// TIA Portal project "ifm-O3D3xx_S7-1200_V16" (V16)

(* hardware
DEVICE "S7-1200 station_1"  S7-1200 Station
   slot 0: "Rack_0"  S7-1200 Rack  Rack  V1.0
   slot 1: "PLC_1"  CPU 1212C AC/DC/Rly  6ES7 212-1BE40-0XB0  V4.4
DEVICE "GSD device_1"  GSD.Device.PN
   slot 0: "Rack"  Rack  V1.0
   slot 0: "O3D3xx"  O3D3XX-PN  O3D3xx  Z1.0
      slot 0: "Standard"  Standard
      slot 1: "Interface"  Interface
         slot 1: "RJ45 10/100 MBit/s"  RJ45 10/100 MBit/s
   slot 1: "450 bytes I_1"  450 bytes I  1.0
      slot 0: "450 bytes I"  450 bytes I
   slot 2: "8 bytes O_1"  8 bytes O  1.0
      slot 0: "8 bytes O"  8 bytes O
DEVICE "HMI_1"  TP700 Comfort
   slot 0: "HMI_1"  TP700 Comfort  6AV2 124-0GC01-0AX0  16.0.0.0
   slot 1: "HMI_RT_1"  TP700 Comfort  6AV2 124-0GC01-0AX0  16.0.0.0
   slot 5: "HMI_1.IE_CP_1"  PROFINET Interface  16.0.0.0
      slot 1: "PROFINET Interface_1"  PROFINET Interface
         slot 1: "Port_1"  Port
         slot 2: "Port_2"  Port
   slot 7: "HMI_1.MPI/DP_CP_1"  MPI/DP Interface  16.0.0.0
DEVICE "GSD device_2"  GSD.Device.PN
   slot 0: "Rack"  Rack  V1.0
   slot 0: "AL1100"  AL1100  AL1100
      slot 0: "AL1100"  AL1100
      slot 1: "X1"  X1
         slot 1: "Port 1"  Port 1
         slot 2: "Port 2"  Port 2
   slot 1: "4 Ports_1"  4 Ports  AL1100
      slot 0: "IO-Link Master"  IO-Link Master
   slot 1: "IO-Link In/Out 32/32 Byte + PQI"  IO-Link In/Out 32/32 Byte + PQI
*)

// ===== PLC "PLC_1"  CPU 1212C AC/DC/Rly =====

VAR_GLOBAL   // PLC tag table "Default tag table"
   "Trigger" AT %M0.0 : Bool;
   "AppNo" AT %MW2 : UInt;
   "GetCounters" AT %M0.1 : Bool;
   "ScrapRate" AT %MD6 : UDInt;
   "Scrap_Alarm" AT %M0.2 : Bool;
   "My_Row_is_OK" AT %M0.3 : Bool;
   "Big Box" AT %M0.4 : Bool;
   "Tag present" AT %I519.2 : Bool;
   "TagValue" AT %IB520 : Byte;
END_VAR

DATA_BLOCK "O3D3xx_Trigger_DB"   // DB1
{ S7_Optimized_Access := 'TRUE' }
AUTHOR : ifm-sy-tl
FAMILY : O3D3xx
VERSION : 1.0
// stored: InstanceOfName O3D3xx_Trigger
"O3D3xx_Trigger"
BEGIN
END_DATA_BLOCK

DATA_BLOCK "O3D3xx_Dimensioning_DB"   // DB2
{ S7_Optimized_Access := 'TRUE' }
AUTHOR : ifm-sy-tl
FAMILY : O3D3xx
VERSION : 1.0
// stored: InstanceOfName O3D3xx_Dimensioning
"O3D3xx_Dimensioning"
BEGIN
END_DATA_BLOCK

DATA_BLOCK "O3D3xx_Completeness_DB"   // DB3
{ S7_Optimized_Access := 'TRUE' }
AUTHOR : ifm-sy-tl
FAMILY : O3D3xx
VERSION : 1.0
// stored: InstanceOfName O3D3xx_Completeness
"O3D3xx_Completeness"
BEGIN
END_DATA_BLOCK

DATA_BLOCK "O3D3xx_GetStatistics_DB"   // DB4
{ S7_Optimized_Access := 'TRUE' }
AUTHOR : ifm-sy-tl
FAMILY : O3D3xx
VERSION : 1.0
// stored: InstanceOfName O3D3xx_GetStatistics
"O3D3xx_GetStatistics"
BEGIN
END_DATA_BLOCK

DATA_BLOCK "ReadData"   // DB5
{ S7_Optimized_Access := 'TRUE' }
VERSION : 0.1
   VAR
      RFIDValue : Byte;
      Object : Struct
         Length : Int;
         Width : Int;
         Height : Int;
      END_STRUCT;
   END_VAR
BEGIN
END_DATA_BLOCK

FUNCTION_BLOCK "O3D3xx_GetStatistics"   // FB8, SCL
TITLE = Get Statistics
{ S7_Optimized_Access := 'TRUE' }
AUTHOR : ifm-sy-tl
FAMILY : O3D3xx
VERSION : 1.1
// executes a "Get Statistics" command and provides the statistics of total, pass and fail readings
   VAR_INPUT
      HW_ID : Hw_Device;   // hardware identifier of the O3D3xx sensor
      Execute : Bool;   // execute Get Statistics command
      TimeoutTime : Time := T#500ms;   // timeout time
   END_VAR
   VAR_OUTPUT
      Done : Bool;   // completed without error
      Busy : Bool;   // command in process
      Error : Bool;   // error occurred
      Status : Word;   // status or error code
      CmdErrorCode : UDInt;   // command error code from O3D3xx sensor
      SysErrorCode : UDInt;   // system error code from O3D3xx sensor
      Total : UDInt;   // total readings
      Pass : UDInt;   // passed readings
      Fail : UDInt;   // failed readings
   END_VAR
   VAR
      tonTimeout : TON_TIME;   // timeout timer of command processing
      diCmdErrorCode : UDInt;   // command error code from O3D3xx sensor
      diSysErrorCode : UDInt;   // system error code from O3D3xx sensor
      wErrorCode : Word;   // current error code of the FB
      iState : Int;   // state of the state machine
      diTotal : UDInt;   // total readings
      diPass : UDInt;   // passed readings
      diFail : UDInt;   // failed readings
   END_VAR
   VAR_TEMP
      Addr : GEOADDR;   // GEO address of the module
      HWModuleID : Hw_Io;   // hardware ID the data module
      DIModuleInAddr : UDInt;   // input address of O3D3xx data
      DIModuleOutAddr : UDInt;   // output address of O3D3xx data
      DIDummy : UDInt;   // dummy
      IModuleInLength : UInt;   // size of data from O3D3xx
      IModuleOutLength : UInt;   // size of data to O3D3xx
      IDummy : UInt;   // dummy
      WCmd : Word;   // command word
      WMirror : Word;   // mirror word
      IResult : Int;   // result of system function
      XDone : Bool;   // task completed
      XError : Bool;   // error detected
      XErrorHW : Bool;   // error hardware assignment
   END_VAR
   VAR CONSTANT
      StateIdle : Int := 16#7000;   // state machine "idle"
      StateSensorRdy : Int := 16#7001;   // state machine "sensor ready"
      StateDeleteError : Int := 16#7002;   // state machine "delete error bit"
      StateGetStatistics : Int := 16#7801;   // state machine "get statistics"
      StateGetError : Int := 16#7601;   // state machine "get error code"
      StateDone : Int := 16#0000;   // state machine "completed"
      StateError : Int := 16#FFFF;   // state machine "error occurred"
   END_VAR
BEGIN
   // Sample program for reading the statistics from an ifm O3D3xx sensor
   // connected to the PLC as Profinet-IO device

   // Function Block Version 1.1.00

   // Description:
   (*
   This FB can be used with an ifm O3D3xx sensor that is connected as Profinet-IO device.
   The core of this FB is to execute a Get Statistics command.
   *)
   // ******************************************************************************************************
   // Disclaimer OF Warranties
   (*
   ifm disclaims to the fullest extent authorized by law any and all warranties,
   whether express or implied, including, without limitation,
   any implied warranties of title, non-infringement, quiet enjoyment,
   integration, merchantability or fitness for a particular purpose.

   Without limitation of the foregoing, ifm expressly does not warrant that:
   (a)  the software will meet your requirements or expectations;
   (b)  the software or the software content will be free of bugs, errors,
        viruses or other defects;
   (c)  any results, output, or data provided through or generated by the software
        will be accurate, up-to-date, complete or reliable;
   (d)  the software will be compatible with third party software;
   (e)  any errors in the software will be corrected


   DEMO SOFTWARE AND TEMPLATES

   Demo software and templates are provided “as is” and “as available”,
   without any warranty of any kind, either express or implied.
   The User acknowledges and agrees to use the software at User’s own risk.
   In no event shall ifm be held liable for any direct, indirect, incidental
   or consequential damages arising out of the use of or inability to use the software.
   User may use the software solely for demonstration purposes
   and to assess the software functionalities and capabilities.


   Software written specifically for Customer

   1. The software created and used is put together by ifm specially to the customer
      using modular software components made by ifm for numerous applications (Standard software modules)
      and adapted to the contractual service required (customer-specific application program).

   2. Upon complete payment of the purchase price for the customer-specific application program,
      ifm transfers the non-exclusive, locally and temporarily unrestricted usage right
      thereof to the customer, without the customer acquiring any rights of any kind
      to the standard software module on which the individual or customer-specific adaptation is based.
      Notwithstanding these provisions, ifm reserves the right to produce and offer
      customer specific software solutions of the same kind for other customers
      based on other terms of reference. In any case ifm retains a simple right of usage
      of the customer–specific solution for internal purposes.

   3. Upon acceptance of the program, User acknowledges and agrees to use the software
      at User’s own risk. User also acknowledges and agrees upon acceptance of the program
      that the software meets the requirements of the specifications agreed upon.
      ifm disclaims any and all warranties, in particular regarding fitness of the software
      for a particular purpose.
   ******************************************************************************************************
   *)

   REGION get addresses and size of O3D3xx data

     // read GEO address of O3D3xx sensor
     #IResult := LOG2GEO(LADDR := #HW_ID, GEOADDR := #Addr);
     #XErrorHW := #IResult <> 0 OR #Addr.AREA <> 1;  // check for error and AREA = PROFINET IO

     #Addr.HWTYPE := 4;  // set hardware type = Module
     #Addr.SUBSLOT := 0;  // set subslot

     REGION  get address and size of INPUT data from O3D3xx
       IF NOT #XErrorHW THEN
         #Addr.SLOT := 1;  // set slot = 1 (slot of INPUT data in O3D3xx configuration)
         #IResult := GEO2LOG(GEOADDR := #Addr, LADDR => #HWModuleID);  // get HW_ID of INPUT data module
         #XErrorHW := #IResult <> 0;  // check for error
       END_IF;
       IF NOT #XErrorHW THEN
         // get IO address of INPUT data
         #IResult := RD_ADDR(LADDR := #HWModuleID,
                             PIADDR => #DIModuleInAddr,
                             PICount => #IModuleInLength,
                             PQADDR => #DIDummy,
                             PQCount => #IDummy);
         #XErrorHW := #IResult <> 0 OR #IDummy <> 0 OR #IModuleInLength <> 64 AND #IModuleInLength <> 450;  // check for error and check size
       END_IF;
     END_REGION get address and size of INPUT data from O3D3xx

     REGION get address and size of OUTPUT data to O3D3xx
       IF NOT #XErrorHW THEN
         #Addr.SLOT := 2;  // set slot = 2 (slot of OUTPUT data in O3D3xx configuration)
         #IResult := GEO2LOG(GEOADDR := #Addr, LADDR => #HWModuleID);  // get HW_ID of OUTPUT data module
         #XErrorHW := #IResult <> 0;  // check for error
       END_IF;
       IF NOT #XErrorHW THEN
         // get IO address of OUTPUT data
         #IResult := RD_ADDR(LADDR := #HWModuleID,
                             PIADDR => #DIDummy,
                             PICount => #IDummy,
                             PQADDR => #DIModuleOutAddr,
                             PQCount => #IModuleOutLength);
         #XErrorHW := #IResult <> 0 OR #IDummy <> 0 OR #IModuleOutLength <> 8;  // check for error and check size
       END_IF;
     END_REGION get address and size of OUTPUT data to O3D3xx

     IF #XErrorHW THEN  // invalid HW_ID
       #wErrorCode := w#16#8100;  // error code for invalid HW_ID
     END_IF;
   END_REGION get addresses and size of O3D3xx data

   REGION read Command Word and Mirror Word of O3D3xx
     IF NOT #XErrorHW THEN
       #WCmd := PEEK_WORD(area := 16#82, dbNumber := 0, byteOffset := UDINT_TO_DINT(IN := #DIModuleOutAddr));
       #WMirror := PEEK_WORD(area := 16#81, dbNumber := 0, byteOffset := UDINT_TO_DINT(IN := #DIModuleInAddr));
     ELSE
       // on error replace values
       #WCmd := w#16#0000;
       #WMirror := w#16#0000;
     END_IF;
   END_REGION read Command Word and Mirror Word of O3D3xx

   REGION reset the Command Bit
     #WCmd := #WCmd AND NOT #WMirror AND w#16#FFFE;  // reset the Command Bit when the Mirror Bit is set
   END_REGION reset the Command Bit

   REGION state machine
     REGION force state machine
       IF #XErrorHW THEN
         // set error state
         #iState := #StateError;
       ELSIF NOT #Execute THEN
         // reset state machine
         #iState := #StateIdle;
       END_IF;
     END_REGION force state machine

     REGION timeout
       CASE #iState OF
         #StateIdle, #StateDone, #StateError:
           #tonTimeout(IN := FALSE,
                       PT := #TimeoutTime);
         ELSE
           #tonTimeout(IN := #WCmd <> w#16#0000,
                       PT := #TimeoutTime);
       END_CASE;
       IF #tonTimeout.Q THEN
         #WCmd := w#16#0000;  // reset all Command Bits
         #wErrorCode := w#16#8205;  // error code for timeout
         #iState := #StateError;
       END_IF;
     END_REGION timeout

     REGION state Idle
       IF #iState = #StateIdle THEN
         #diCmdErrorCode := 0;  // initialize error codes
         #diSysErrorCode := 0;
         IF #Execute THEN
           // input EXECUTE active
           #iState := #StateSensorRdy;
         END_IF;  // input EXECUTE active
       END_IF;
     END_REGION state Idle

     REGION state Sensor Ready
       IF #iState = #StateSensorRdy THEN
         IF #WCmd <> w#16#0000 THEN
           // any Command Bit is set
           #wErrorCode := w#16#8301;  // error code for other command active
           #iState := #StateError;
         ELSIF (#WMirror AND w#16#FFFE) = w#16#0000 THEN
           // all Mirror Bits reset
           IF #WMirror.%X0 THEN
             // Error bit is set
             #iState := #StateDeleteError;
           ELSE
             // no previous error
             #iState := #StateGetStatistics;
           END_IF;  // no previous error
         END_IF;  // all Mirror Bits reset
       END_IF;
     END_REGION state Sensor Ready

     REGION state Delete Error Bit
       IF #iState = #StateDeleteError THEN
         IF NOT #WMirror.%X6 THEN
           // set Get Error command bit
           #WCmd.%X6 := TRUE;
         ELSE
           // Get Error command finished
           IF #WMirror.%X0 THEN
             // Error bit still set
             #wErrorCode := w#16#8001;  // error code for error remains active
             #iState := #StateError;
           ELSE
             // Error bit is reset
             #iState := #StateGetStatistics;
           END_IF;  // Error bit is reset
         END_IF;  // Get Error command finished
       END_IF;
     END_REGION state Delete Error Bit

     REGION state Get Statistics
       IF #iState = #StateGetStatistics THEN
         IF NOT #WMirror.%X8 THEN
           // set Get Statistics command bit
           #WCmd.%X8 := TRUE;
         ELSE
           // Get Statistics command finished
           IF #WMirror.%X0 THEN
             // error occurred
             #iState := #StateGetError;
           ELSE
             // no error
             // read reported statistics
             #diTotal := DWORD_TO_UDINT(PEEK_DWORD(area := 16#81, dbNumber := 0, byteOffset := UDINT_TO_DINT(IN := #DIModuleInAddr + 8)));
             #diPass := DWORD_TO_UDINT(PEEK_DWORD(area := 16#81, dbNumber := 0, byteOffset := UDINT_TO_DINT(IN := #DIModuleInAddr + 12)));
             #diFail := DWORD_TO_UDINT(PEEK_DWORD(area := 16#81, dbNumber := 0, byteOffset := UDINT_TO_DINT(IN := #DIModuleInAddr + 16)));
             #iState := #StateDone;
           END_IF;  // no error
         END_IF;  // Get Statistics command finished
       END_IF;
     END_REGION state Get Statistics

     REGION state Get Error Code
       IF #iState = #StateGetError THEN
         IF NOT #WMirror.%X6 THEN
           // set Get Error command bit
           #WCmd.%X6 := TRUE;
         ELSE
           // Get Error command finished
           #wErrorCode := w#16#8000;  // error code for sensor error
           // read reported command error and system error codes
           #diCmdErrorCode := DWORD_TO_UDINT(PEEK_DWORD(area := 16#81, dbNumber := 0, byteOffset := UDINT_TO_DINT(IN := #DIModuleInAddr + 8)));
           #diSysErrorCode := DWORD_TO_UDINT(PEEK_DWORD(area := 16#81, dbNumber := 0, byteOffset := UDINT_TO_DINT(IN := #DIModuleInAddr + 12)));
           #iState := #StateError;
         END_IF;  // Get Error command finished
       END_IF;
     END_REGION state Get Error Code 
   END_REGION state machine

   REGION set OUTPUTS to the O3D3xx sensor
     IF NOT #XErrorHW THEN
       // hardware is accessible
       POKE(area := 16#82,
            dbNumber := 0,
            byteOffset := UDINT_TO_DINT(#DIModuleOutAddr),
            value := #WCmd);
     END_IF;
   END_REGION set OUTPUTS to the O3D3xx sensor

   REGION set FB outputs
     #XDone := #iState = #StateDone;
     #XError := #iState = #StateError;

     #Done := #XDone;  // show command completeed
     #Busy := #Execute AND NOT #XDone AND NOT #XError;  // show that the command processing is active
     #Error := #XError;  // show that an error occurred
     IF #XError THEN
       // on error show error codes
       #Status := #wErrorCode;
       #CmdErrorCode := #diCmdErrorCode;
       #SysErrorCode := #diSysErrorCode;
     ELSE
       // in normal operation
       #Status := INT_TO_WORD(#iState);  // show active state
       #CmdErrorCode := 0;  // show no error codes
       #SysErrorCode := 0;
     END_IF;
     IF #XDone THEN
       // when command is completed, show statistics
       #Total := #diTotal;
       #Pass := #diPass;
       #Fail := #diFail;
     ELSE
       // show initial values
       #Total := 0;
       #Pass := 0;
       #Fail := 0;
     END_IF;  // schow initial values
   END_REGION set FB outputs
END_FUNCTION_BLOCK

FUNCTION_BLOCK "O3D3xx_Trigger"   // FB13, SCL
TITLE = Trigger
{ S7_Optimized_Access := 'TRUE' }
AUTHOR : ifm-sy-tl
FAMILY : O3D3xx
VERSION : 1.0
// executes a "Synchronous Trigger" command with the option to activate a specific application in the sensor before triggering the sensor
   VAR_INPUT
      HW_ID : Hw_Device;   // hardware identifier of the O3D3xx sensor
      Execute : Bool;   // trigger the O3D3xx sensor
      AppNo : UInt := 0;   // application No. to activate [1..32]
      TimeoutTime : Time := T#2000ms;   // timeout time
   END_VAR
   VAR_OUTPUT
      Done : Bool;   // completed without error
      Busy : Bool;   // command in process
      Error : Bool;   // error occurred
      Status : Word;   // status or error code
      CmdErrorCode : UDInt;   // command error code from O3D3xx sensor
      SysErrorCode : UDInt;   // system error code from O3D3xx sensor
   END_VAR
   VAR
      tonTimeout : TON_TIME;   // timeout timer of command processing
      diCmdErrorCode : UDInt;   // command error code from O3D3xx sensor
      diSysErrorCode : UDInt;   // system error code from O3D3xx sensor
      wErrorCode : Word;   // current error code of the FB
      iState : Int;   // state of the state machine
      iAppNo : UInt;   // application No. to activate
   END_VAR
   VAR_TEMP
      Addr : GEOADDR;   // GEO address of the module
      HWModuleID : Hw_Io;   // hardware ID the data module
      DIModuleInAddr : UDInt;   // input address of O3D3xx data
      DIModuleOutAddr : UDInt;   // output address of O3D3xx data
      DIDummy : UDInt;   // dummy
      IModuleInLength : UInt;   // size of data from O3D3xx
      IModuleOutLength : UInt;   // size of data to O3D3xx
      IDummy : UInt;   // dummy
      WCmd : Word;   // command word
      WMirror : Word;   // mirror word
      IResult : Int;   // result of system function
      XDone : Bool;   // task completed
      XError : Bool;   // error detected
      XErrorHW : Bool;   // error hardware assignment
   END_VAR
   VAR CONSTANT
      StateIdle : Int := 16#7000;   // state machine "idle"
      StateSensorRdy : Int := 16#7001;   // state machine "sensor ready"
      StateDeleteError : Int := 16#7002;   // state machine "delete error bit"
      StateActivateApp : Int := 16#7901;   // state machine "activate app"
      StateTrigger : Int := 16#7D01;   // state machine "trigger"
      StateGetError : Int := 16#7601;   // state machine "get error code"
      StateDone : Int := 16#0000;   // state machine "completed"
      StateError : Int := 16#FFFF;   // state machine "error occurred"
   END_VAR
BEGIN
   // Sample program to trigger an ifm O3D3xx sensor
   // connected to the PLC as Profinet-IO device

   // Function Block Version 1.0.00

   // Description:
   (*
   This FB can be used with an ifm O3D3xx sensor that is connected as Profinet-IO device.
   The core of this FB is to execute a Synchronous Trigger command.
   If the assigned value at the parameter AppNo > 0 the FB activates the assigned application in the sensor
   before it executes the trigger command.
   *)
   // ******************************************************************************************************
   // Disclaimer OF Warranties
   (*
   ifm disclaims to the fullest extent authorized by law any and all warranties,
   whether express or implied, including, without limitation,
   any implied warranties of title, non-infringement, quiet enjoyment,
   integration, merchantability or fitness for a particular purpose.

   Without limitation of the foregoing, ifm expressly does not warrant that:
   (a)  the software will meet your requirements or expectations;
   (b)  the software or the software content will be free of bugs, errors,
        viruses or other defects;
   (c)  any results, output, or data provided through or generated by the software
        will be accurate, up-to-date, complete or reliable;
   (d)  the software will be compatible with third party software;
   (e)  any errors in the software will be corrected


   DEMO SOFTWARE AND TEMPLATES

   Demo software and templates are provided “as is” and “as available”,
   without any warranty of any kind, either express or implied.
   The User acknowledges and agrees to use the software at User’s own risk.
   In no event shall ifm be held liable for any direct, indirect, incidental
   or consequential damages arising out of the use of or inability to use the software.
   User may use the software solely for demonstration purposes
   and to assess the software functionalities and capabilities.


   Software written specifically for Customer

   1. The software created and used is put together by ifm specially to the customer
      using modular software components made by ifm for numerous applications (Standard software modules)
      and adapted to the contractual service required (customer-specific application program).

   2. Upon complete payment of the purchase price for the customer-specific application program,
      ifm transfers the non-exclusive, locally and temporarily unrestricted usage right
      thereof to the customer, without the customer acquiring any rights of any kind
      to the standard software module on which the individual or customer-specific adaptation is based.
      Notwithstanding these provisions, ifm reserves the right to produce and offer
      customer specific software solutions of the same kind for other customers
      based on other terms of reference. In any case ifm retains a simple right of usage
      of the customer–specific solution for internal purposes.

   3. Upon acceptance of the program, User acknowledges and agrees to use the software
      at User’s own risk. User also acknowledges and agrees upon acceptance of the program
      that the software meets the requirements of the specifications agreed upon.
      ifm disclaims any and all warranties, in particular regarding fitness of the software
      for a particular purpose.
   ******************************************************************************************************
   *)

   REGION get addresses and size of O3D3xx data

     // read GEO address of O3D3xx sensor
     #IResult := LOG2GEO(LADDR := #HW_ID, GEOADDR := #Addr);
     #XErrorHW := #IResult <> 0 OR #Addr.AREA <> 1;  // check for error and AREA = PROFINET IO

     #Addr.HWTYPE := 4;  // set hardware type = Module
     #Addr.SUBSLOT := 0;  // set subslot

     REGION  get address and size of INPUT data from O3D3xx
       IF NOT #XErrorHW THEN
         #Addr.SLOT := 1;  // set slot = 1 (slot of INPUT data in O3D3xx configuration)
         #IResult := GEO2LOG(GEOADDR := #Addr, LADDR => #HWModuleID);  // get HW_ID of INPUT data module
         #XErrorHW := #IResult <> 0;  // check for error
       END_IF;
       IF NOT #XErrorHW THEN
         // get IO address of INPUT data
         #IResult := RD_ADDR(LADDR := #HWModuleID,
                             PIADDR => #DIModuleInAddr,
                             PICount => #IModuleInLength,
                             PQADDR => #DIDummy,
                             PQCount => #IDummy);
         #XErrorHW := #IResult <> 0 OR #IDummy <> 0 OR #IModuleInLength <> 64 AND #IModuleInLength <> 450;  // check for error and check size
       END_IF;
     END_REGION get address and size of INPUT data from O3D3xx

     REGION get address and size of OUTPUT data to O3D3xx
       IF NOT #XErrorHW THEN
         #Addr.SLOT := 2;  // set slot = 2 (slot of OUTPUT data in O3D3xx configuration)
         #IResult := GEO2LOG(GEOADDR := #Addr, LADDR => #HWModuleID);  // get HW_ID of OUTPUT data module
         #XErrorHW := #IResult <> 0;  // check for error
       END_IF;
       IF NOT #XErrorHW THEN
         // get IO address of OUTPUT data
         #IResult := RD_ADDR(LADDR := #HWModuleID,
                             PIADDR => #DIDummy,
                             PICount => #IDummy,
                             PQADDR => #DIModuleOutAddr,
                             PQCount => #IModuleOutLength);
         #XErrorHW := #IResult <> 0 OR #IDummy <> 0 OR #IModuleOutLength <> 8;  // check for error and check size
       END_IF;
     END_REGION get address and size of OUTPUT data to O3D3xx

     IF #XErrorHW THEN  // invalid HW_ID
       #wErrorCode := w#16#8100;  // error code for invalid HW_ID
     END_IF;
   END_REGION get addresses and size of O3D3xx data

   REGION read Command Word and Mirror Word of O3D3xx
     IF NOT #XErrorHW THEN
       #WCmd := PEEK_WORD(area := 16#82, dbNumber := 0, byteOffset := UDINT_TO_DINT(IN := #DIModuleOutAddr));
       #WMirror := PEEK_WORD(area := 16#81, dbNumber := 0, byteOffset := UDINT_TO_DINT(IN := #DIModuleInAddr));
     ELSE
       // on error replace values
       #WCmd := w#16#0000;
       #WMirror := w#16#0000;
     END_IF;
   END_REGION read Command Word and Mirror Word of O3D3xx

   REGION reset the Command Bit
     #WCmd := #WCmd AND NOT #WMirror AND w#16#FFFE;  // reset the Command Bit when the Mirror Bit is set
   END_REGION reset the Command Bit

   REGION state machine
     REGION force state machine
       IF #XErrorHW THEN
         // set error state
         #iState := #StateError;
       ELSIF NOT #Execute THEN
         // reset state machine
         #iState := #StateIdle;
       END_IF;
     END_REGION force state machine

     REGION timeout
       CASE #iState OF
         #StateIdle, #StateDone, #StateError:
           #tonTimeout(IN := FALSE,
                       PT := #TimeoutTime);
         ELSE
           #tonTimeout(IN := #WCmd <> w#16#0000,
                       PT := #TimeoutTime);
       END_CASE;
       IF #tonTimeout.Q THEN
         #WCmd := w#16#0000;  // reset all Command Bits
         #wErrorCode := w#16#8205;  // error code for timeout
         #iState := #StateError;
       END_IF;
     END_REGION timeout

     REGION state Idle
       IF #iState = #StateIdle THEN
         #diCmdErrorCode := 0;  // initialize error codes
         #diSysErrorCode := 0;
         IF #Execute THEN
           // input EXECUTE active
           IF #AppNo > 32 THEN
             // Application Number is invalid
             #wErrorCode := w#16#8302;  // set error code
             #iState := #StateError;
           ELSE
             // Application Number is valid
             #iAppNo := #AppNo;  // store parameter value
             #iState := #StateSensorRdy;
           END_IF;  // Application Number is valid
         END_IF;  // input EXECUTE active
       END_IF;
     END_REGION state Idle

     REGION state Sensor Ready
       IF #iState = #StateSensorRdy THEN
         IF #WCmd <> w#16#0000 THEN
           // any Command Bit is set
           #wErrorCode := w#16#8301;  // error code for other command active
           #iState := #StateError;
         ELSIF (#WMirror AND w#16#FFFE) = w#16#0000 THEN
           // all Mirror Bits reset
           IF #WMirror.%X0 THEN
             // Error bit is set
             #iState := #StateDeleteError;
           ELSIF #iAppNo = 0 THEN
             // trigger only
             #iState := #StateTrigger;
           ELSE
             // activate application before trigger
             #iState := #StateActivateApp;
           END_IF;  // activate application before trigger
         END_IF;  // all Mirror Bits reset
       END_IF;
     END_REGION state Sensor Ready

     REGION state Delete Error Bit
       IF #iState = #StateDeleteError THEN
         IF NOT #WMirror.%X6 THEN
           // set Get Error command bit
           #WCmd.%X6 := TRUE;
         ELSE
           // Get Error command finished
           IF #WMirror.%X0 THEN
             // Error bit still set
             #wErrorCode := w#16#8001;  // error code for error remains active
             #iState := #StateError;
           ELSIF #iAppNo = 0 THEN
             // trigger only
             #iState := #StateTrigger;
           ELSE
             // activate application before trigger
             #iState := #StateActivateApp;
           END_IF;  // activate application before trigger
         END_IF;  // Get Error command finished
       END_IF;
     END_REGION state Delete Error Bit

     REGION state Activate Application
       IF #iState = #StateActivateApp THEN
         IF NOT #WMirror.%X9 THEN
             // set Activate Application command bit and command parameter
           #WCmd.%X9 := TRUE;
           POKE(area := 16#82,
                dbNumber := 0,
                byteOffset := UDINT_TO_DINT(IN := #DIModuleOutAddr + 2),
                value := w#16#0000);
           POKE(area := 16#82,
                dbNumber := 0,
                byteOffset := UDINT_TO_DINT(IN := #DIModuleOutAddr + 4),
                value := w#16#0000);
           POKE(area := 16#82,
                dbNumber := 0,
                byteOffset := UDINT_TO_DINT(IN := #DIModuleOutAddr + 6),
                value := UINT_TO_WORD(#iAppNo));
         ELSE
           // Activate Application command finished
           IF #WMirror.%X0 THEN
             // error occurred
             #iState := #StateGetError;
           ELSE
             // no error
             #iState := #StateTrigger;
           END_IF;  // no error
         END_IF;  // Activate Application command finished
       END_IF;
     END_REGION state Activate Application

     REGION state Trigger
       IF #iState = #StateTrigger THEN
         IF NOT #WMirror.%X13 THEN
           // set Trigger command bit
           #WCmd.%X13 := TRUE;
         ELSE
           // Trigger command finished
           IF #WMirror.%X0 THEN
             // error occurred
             #iState := #StateGetError;
           ELSE
             // no error
             #iState := #StateDone;
           END_IF;  // no error
         END_IF;  // Trigger command finished
       END_IF;
     END_REGION state Trigger

     REGION state Get Error Code
       IF #iState = #StateGetError THEN
         IF NOT #WMirror.%X6 THEN
           // set Get Error command bit
           #WCmd.%X6 := TRUE;
         ELSE
           // Get Error command finished
           #wErrorCode := w#16#8000;  // error code for sensor error
           // read reported command error and system error codes
           #diCmdErrorCode := DWORD_TO_UDINT(PEEK_DWORD(area := 16#81, dbNumber := 0, byteOffset := UDINT_TO_DINT(IN := #DIModuleInAddr + 8)));
           #diSysErrorCode := DWORD_TO_UDINT(PEEK_DWORD(area := 16#81, dbNumber := 0, byteOffset := UDINT_TO_DINT(IN := #DIModuleInAddr + 12)));
           #iState := #StateError;
         END_IF;  // Get Error command finished
       END_IF;
     END_REGION state Get Error Code 
   END_REGION state machine

   REGION set OUTPUTS to the O3D3xx sensor
     IF NOT #XErrorHW THEN
       // hardware is accessible
       POKE(area := 16#82,
            dbNumber := 0,
            byteOffset := UDINT_TO_DINT(#DIModuleOutAddr),
            value := #WCmd);
     END_IF;
   END_REGION set OUTPUTS to the O3D3xx sensor

   REGION set FB outputs
     #XDone := #iState = #StateDone;
     #XError := #iState = #StateError;

     #Done := #XDone;  // show command completeed
     #Busy := #Execute AND NOT #XDone AND NOT #XError;  // show that the command processing is active
     #Error := #XError;  // show that an error occurred
     IF #XError THEN
       // on error show error codes
       #Status := #wErrorCode;
       #CmdErrorCode := #diCmdErrorCode;
       #SysErrorCode := #diSysErrorCode;
     ELSE
       // in normal operation
       #Status := INT_TO_WORD(#iState);  // show active state
       #CmdErrorCode := 0;  // show no error codes
       #SysErrorCode := 0;
     END_IF;
   END_REGION set FB outputs
END_FUNCTION_BLOCK

FUNCTION_BLOCK "O3D3xx_Dimensioning"   // FB23, SCL
TITLE = Dimensioning Wizard Result
{ S7_Optimized_Access := 'TRUE' }
AUTHOR : ifm-sy-tl
FAMILY : O3D3xx
VERSION : 1.0
// monitors the input data from the sensor and interpretes trigger result data according to the data output definition of the “Dimensioning” application wizard of the ifmVisionAssistant software V1.8
   VAR_INPUT
      HW_ID : Hw_Device;   // hardware identifier of the O3D3xx sensor
   END_VAR
   VAR_OUTPUT
      ErrorCodeFB : Word;   // error code of the function block
      NewData : Bool;   // new data
      ObjectFound : Bool;   // object found
      Width : Int;   // width of object
      Height : Int;   // height of object
      Length : Int;   // length of object
      PosX : Int;   // x-coordinate of object
      PosY : Int;   // y-coordinate of object
      PosZ : Int;   // z-coordinate of object
      Angle : Int;   // angle of rotation of object
      QualityW : Int;   // quality of width value
      QualityH : Int;   // quality of height value
      QualityL : Int;   // quality of length value
   END_VAR
   VAR
      iprevMsgCounter : UInt;   // previous message counter value
      xprevMirrorbit : Bool;   // previous state of the Mirror Bit
   END_VAR
   VAR_TEMP
      Addr : GEOADDR;   // GEO address of the module
      HWModuleID : Hw_Io;   // hardware ID the data module
      DIModuleInAddr : UDInt;   // input address of O3D3xx data
      DIDummy : UDInt;   // dummy
      IModuleInLength : UInt;   // size of data from O3D3xx
      IDummy : UInt;   // dummy
      WMsgID : Word;   // current message ID
      IMsgCounter : UInt;   // current message counter
      IResult : Int;   // result of system function
      XTriggerMirrorbit : Bool;   // Mirror Bit of Trigger command
      XreMirrorbit : Bool;   // rising edge of Mirror Bit
      XreNewAsyncResult : Bool;   // new asynchronous result message
      XErrorHW : Bool;   // error hardware assignment
   END_VAR
BEGIN
   // Sample program for detecting and interpreting result data from an ifm O3D3xx sensor
   // connected to the PLC as Profinet-IO device

   // “Dimensioning” application wizard
   // Function Block Version 1.0.00

   // Description:
   (*
   This FB can be used with an ifm O3D3xx sensor that is connected as Profinet-IO device.
   It monitors the input data from the O3D3xx sensor.
   If the FB identifies a trigger result, it interprets the data according to the data output definition of the
   “Dimensioning of rectangular objects” application wizard of the ifmVisionAssistant software V1.8.
   The signal "NewData" rises for one PLC cycle. The data remain in the outputs until the next data are received.
   *)
   // ******************************************************************************************************
   // Disclaimer OF Warranties
   (*
   ifm disclaims to the fullest extent authorized by law any and all warranties,
   whether express or implied, including, without limitation,
   any implied warranties of title, non-infringement, quiet enjoyment,
   integration, merchantability or fitness for a particular purpose.

   Without limitation of the foregoing, ifm expressly does not warrant that:
   (a)  the software will meet your requirements or expectations;
   (b)  the software or the software content will be free of bugs, errors,
        viruses or other defects;
   (c)  any results, output, or data provided through or generated by the software
        will be accurate, up-to-date, complete or reliable;
   (d)  the software will be compatible with third party software;
   (e)  any errors in the software will be corrected


   DEMO SOFTWARE AND TEMPLATES

   Demo software and templates are provided “as is” and “as available”,
   without any warranty of any kind, either express or implied.
   The User acknowledges and agrees to use the software at User’s own risk.
   In no event shall ifm be held liable for any direct, indirect, incidental
   or consequential damages arising out of the use of or inability to use the software.
   User may use the software solely for demonstration purposes
   and to assess the software functionalities and capabilities.


   Software written specifically for Customer

   1. The software created and used is put together by ifm specially to the customer
      using modular software components made by ifm for numerous applications (Standard software modules)
      and adapted to the contractual service required (customer-specific application program).

   2. Upon complete payment of the purchase price for the customer-specific application program,
      ifm transfers the non-exclusive, locally and temporarily unrestricted usage right
      thereof to the customer, without the customer acquiring any rights of any kind
      to the standard software module on which the individual or customer-specific adaptation is based.
      Notwithstanding these provisions, ifm reserves the right to produce and offer
      customer specific software solutions of the same kind for other customers
      based on other terms of reference. In any case ifm retains a simple right of usage
      of the customer–specific solution for internal purposes.

   3. Upon acceptance of the program, User acknowledges and agrees to use the software
      at User’s own risk. User also acknowledges and agrees upon acceptance of the program
      that the software meets the requirements of the specifications agreed upon.
      ifm disclaims any and all warranties, in particular regarding fitness of the software
      for a particular purpose.
   ******************************************************************************************************
   *)

   REGION get address and size of INPUT data from O3D3xx    
     #IResult := LOG2GEO(LADDR := #HW_ID, GEOADDR := #Addr);  // read GEO address of O3D3xx sensor
     #XErrorHW := #IResult <> 0 OR #Addr.AREA <> 1;  // check for error and AREA = PROFINET IO
     IF NOT #XErrorHW THEN
       #Addr.HWTYPE := 4;  // set hardware type = Module
       #Addr.SLOT := 1;  // set slot = 1 (slot of INPUT data in O3D3xx configuration)
       #Addr.SUBSLOT := 0;  // set subslot
       #IResult := GEO2LOG(GEOADDR := #Addr, LADDR => #HWModuleID);  // get HW_ID of INPUT data module
       #XErrorHW := #IResult <> 0;  // check for error
     END_IF;
     IF NOT #XErrorHW THEN
       // get IO address of INPUT data
       #IResult := RD_ADDR(LADDR := #HWModuleID,
                           PIADDR => #DIModuleInAddr,
                           PICount => #IModuleInLength,
                           PQADDR => #DIDummy,
                           PQCount => #IDummy);
       #XErrorHW := #IResult <> 0 OR #IDummy <> 0 OR #IModuleInLength <> 64 AND #IModuleInLength <> 450;  // check for error and check size
     END_IF;
   END_REGION get address and size of INPUT data from O3D3xx

   REGION read input data header of O3D3xx
     IF NOT #XErrorHW THEN
       #XTriggerMirrorbit := PEEK_BOOL(area := 16#81, dbNumber := 0, byteOffset := UDINT_TO_DINT(IN := #DIModuleInAddr), bitOffset := 5);
       #WMsgID := PEEK_WORD(area := 16#81, dbNumber := 0, byteOffset := UDINT_TO_DINT(IN := #DIModuleInAddr + 2));
       #IMsgCounter := WORD_TO_UINT(PEEK_WORD(area := 16#81, dbNumber := 0, byteOffset := UDINT_TO_DINT(IN := #DIModuleInAddr + 4)));

       REGION check for new result
         // check for new synchronous result
         #XreMirrorbit := #XTriggerMirrorbit AND NOT #xprevMirrorbit;  // detect rising edge of the Mirror Bit
         #xprevMirrorbit := #XTriggerMirrorbit;  // store current state to detect the change

         //  check for new asynchronous result
         #XreNewAsyncResult := #IMsgCounter <> #iprevMsgCounter AND #WMsgID = w#16#0001;  // new asynchronous result received
         #iprevMsgCounter := #IMsgCounter;  // store current value to detect the change
       END_REGION check for new result
     ELSE
       // on error replace values
       #XreMirrorbit := FALSE;
       #XreNewAsyncResult := FALSE;
     END_IF;  // on error replace values
   END_REGION read input data header of O3D3xx

   REGION set FB outputs
     IF #XErrorHW THEN  // invalid HW_ID
       #ErrorCodeFB := w#16#8100;  // error code for invalid HW_ID
     ELSE
       #ErrorCodeFB := w#16#0000;
     END_IF;
     #NewData := #XreMirrorbit OR #XreNewAsyncResult;  // new trigger response data
     IF #XreMirrorbit OR #XreNewAsyncResult THEN
       // transfer data into outputs
       #ObjectFound := w#16#0001 = PEEK_WORD(area := 16#81, dbNumber := 0, byteOffset := UDINT_TO_DINT(IN := #DIModuleInAddr + 12));
       #Width := WORD_TO_INT(PEEK_WORD(area := 16#81, dbNumber := 0, byteOffset := UDINT_TO_DINT(IN := #DIModuleInAddr + 14)));
       #Height := WORD_TO_INT(PEEK_WORD(area := 16#81, dbNumber := 0, byteOffset := UDINT_TO_DINT(IN := #DIModuleInAddr + 16)));
       #Length := WORD_TO_INT(PEEK_WORD(area := 16#81, dbNumber := 0, byteOffset := UDINT_TO_DINT(IN := #DIModuleInAddr + 18)));
       #PosX := WORD_TO_INT(PEEK_WORD(area := 16#81, dbNumber := 0, byteOffset := UDINT_TO_DINT(IN := #DIModuleInAddr + 20)));
       #PosY := WORD_TO_INT(PEEK_WORD(area := 16#81, dbNumber := 0, byteOffset := UDINT_TO_DINT(IN := #DIModuleInAddr + 22)));
       #PosZ := WORD_TO_INT(PEEK_WORD(area := 16#81, dbNumber := 0, byteOffset := UDINT_TO_DINT(IN := #DIModuleInAddr + 24)));
       #Angle := WORD_TO_INT(PEEK_WORD(area := 16#81, dbNumber := 0, byteOffset := UDINT_TO_DINT(IN := #DIModuleInAddr + 26)));
       #QualityW := WORD_TO_INT(PEEK_WORD(area := 16#81, dbNumber := 0, byteOffset := UDINT_TO_DINT(IN := #DIModuleInAddr + 28)));
       #QualityH := WORD_TO_INT(PEEK_WORD(area := 16#81, dbNumber := 0, byteOffset := UDINT_TO_DINT(IN := #DIModuleInAddr + 30)));
       #QualityL := WORD_TO_INT(PEEK_WORD(area := 16#81, dbNumber := 0, byteOffset := UDINT_TO_DINT(IN := #DIModuleInAddr + 32)));
     END_IF;  // transfer data into outputs
   END_REGION set FB outputs
END_FUNCTION_BLOCK

FUNCTION_BLOCK "O3D3xx_Completeness"   // FB25, SCL
TITLE = Completeness Wizard Result
{ S7_Optimized_Access := 'TRUE' }
AUTHOR : ifm-sy-tl
FAMILY : O3D3xx
VERSION : 1.0
// monitors the input data from the sensor and interpretes trigger result data according to the data output definition of the “Completeness” application wizard of the ifmVisionAssistant software V1.8
   VAR_INPUT
      HW_ID : Hw_Device;   // hardware identifier of the O3D3xx sensor
      Tracking : Bool;   // anchor tracking enabled in the O3D3xx application
   END_VAR
   VAR_OUTPUT
      ErrorCodeFB : Word;   // error code of the function block
      NewData : Bool;   // new data
      TrackingOK : Bool;   // anchor tracking successful
      AllROIsGood : Bool;   // result of all ROIs = OK
      ROI : Array[0..63] of Struct   // ROI results
         Status : Int;   // ROI status
         Value : Int;   // ROI value [mm]
      END_STRUCT;
   END_VAR
   VAR
      iprevMsgCounter : UInt;   // previous message counter value
      xprevMirrorbit : Bool;   // previous state of the Mirror Bit
   END_VAR
   VAR_TEMP
      Addr : GEOADDR;   // GEO address of the module
      HWModuleID : Hw_Io;   // hardware ID the data module
      DIModuleInAddr : UDInt;   // input address of O3D3xx data
      DIDummy : UDInt;   // dummy
      IModuleInLength : UInt;   // size of data from O3D3xx
      IDummy : UInt;   // dummy
      WMsgID : Word;   // current message ID
      IMsgCounter : UInt;   // current message counter
      IResult : Int;   // result of system function
      DIRdAddr : DInt;   // read address
      DILastRdAddr : DInt;   // start address of last dataset
      IID : Int;   // ROI ID
      XTriggerMirrorbit : Bool;   // Mirror Bit of Trigger command
      XreMirrorbit : Bool;   // rising edge of Mirror Bit
      XreNewAsyncResult : Bool;   // new asynchronous result message
      XErrorHW : Bool;   // error hardware assignment
   END_VAR
BEGIN
   // Sample program for detecting and interpreting result data from an ifm O3D3xx sensor
   // connected to the PLC as Profinet-IO device

   // “Completeness” application wizard
   // Function Block Version 1.0.00

   // Description:
   (*
   This FB can be used with an ifm O3D3xx sensor that is connected as Profinet-IO device.
   It monitors the input data from the O3D3xx sensor.
   If the FB identifies a trigger result, it interprets the data according to the data output definition of the
   “Completeness” application wizard of the ifmVisionAssistant software V1.8.
   The signal "NewData" rises for one PLC cycle. The data remain in the outputs until the next data are received.
   *)
   // ******************************************************************************************************
   // Disclaimer OF Warranties
   (*
   ifm disclaims to the fullest extent authorized by law any and all warranties,
   whether express or implied, including, without limitation,
   any implied warranties of title, non-infringement, quiet enjoyment,
   integration, merchantability or fitness for a particular purpose.

   Without limitation of the foregoing, ifm expressly does not warrant that:
   (a)  the software will meet your requirements or expectations;
   (b)  the software or the software content will be free of bugs, errors,
        viruses or other defects;
   (c)  any results, output, or data provided through or generated by the software
        will be accurate, up-to-date, complete or reliable;
   (d)  the software will be compatible with third party software;
   (e)  any errors in the software will be corrected


   DEMO SOFTWARE AND TEMPLATES

   Demo software and templates are provided “as is” and “as available”,
   without any warranty of any kind, either express or implied.
   The User acknowledges and agrees to use the software at User’s own risk.
   In no event shall ifm be held liable for any direct, indirect, incidental
   or consequential damages arising out of the use of or inability to use the software.
   User may use the software solely for demonstration purposes
   and to assess the software functionalities and capabilities.


   Software written specifically for Customer

   1. The software created and used is put together by ifm specially to the customer
      using modular software components made by ifm for numerous applications (Standard software modules)
      and adapted to the contractual service required (customer-specific application program).

   2. Upon complete payment of the purchase price for the customer-specific application program,
      ifm transfers the non-exclusive, locally and temporarily unrestricted usage right
      thereof to the customer, without the customer acquiring any rights of any kind
      to the standard software module on which the individual or customer-specific adaptation is based.
      Notwithstanding these provisions, ifm reserves the right to produce and offer
      customer specific software solutions of the same kind for other customers
      based on other terms of reference. In any case ifm retains a simple right of usage
      of the customer–specific solution for internal purposes.

   3. Upon acceptance of the program, User acknowledges and agrees to use the software
      at User’s own risk. User also acknowledges and agrees upon acceptance of the program
      that the software meets the requirements of the specifications agreed upon.
      ifm disclaims any and all warranties, in particular regarding fitness of the software
      for a particular purpose.
   ******************************************************************************************************
   *)

   REGION get address and size of INPUT data from O3D3xx    
     #IResult := LOG2GEO(LADDR := #HW_ID, GEOADDR := #Addr);  // read GEO address of O3D3xx sensor
     #XErrorHW := #IResult <> 0 OR #Addr.AREA <> 1;  // check for error and AREA = PROFINET IO
     IF NOT #XErrorHW THEN
       #Addr.HWTYPE := 4;  // set hardware type = Module
       #Addr.SLOT := 1;  // set slot = 1 (slot of INPUT data in O3D3xx configuration)
       #Addr.SUBSLOT := 0;  // set subslot
       #IResult := GEO2LOG(GEOADDR := #Addr, LADDR => #HWModuleID);  // get HW_ID of INPUT data module
       #XErrorHW := #IResult <> 0;  // check for error
     END_IF;
     IF NOT #XErrorHW THEN
       // get IO address of INPUT data
       #IResult := RD_ADDR(LADDR := #HWModuleID,
                           PIADDR => #DIModuleInAddr,
                           PICount => #IModuleInLength,
                           PQADDR => #DIDummy,
                           PQCount => #IDummy);
       #XErrorHW := #IResult <> 0 OR #IDummy <> 0 OR #IModuleInLength <> 64 AND #IModuleInLength <> 450;  // check for error and check size
     END_IF;
   END_REGION get address and size of INPUT data from O3D3xx

   REGION read input data header of O3D3xx
     IF NOT #XErrorHW THEN
       #XTriggerMirrorbit := PEEK_BOOL(area := 16#81, dbNumber := 0, byteOffset := UDINT_TO_DINT(IN := #DIModuleInAddr), bitOffset := 5);
       #WMsgID := PEEK_WORD(area := 16#81, dbNumber := 0, byteOffset := UDINT_TO_DINT(IN := #DIModuleInAddr + 2));
       #IMsgCounter := WORD_TO_UINT(PEEK_WORD(area := 16#81, dbNumber := 0, byteOffset := UDINT_TO_DINT(IN := #DIModuleInAddr + 4)));

       REGION check for new result
         // check for new synchronous result
         #XreMirrorbit := #XTriggerMirrorbit AND NOT #xprevMirrorbit;  // detect rising edge of the Mirror Bit
         #xprevMirrorbit := #XTriggerMirrorbit;  // store current state to detect the change

         //  check for new asynchronous result
         #XreNewAsyncResult := #IMsgCounter <> #iprevMsgCounter AND #WMsgID = w#16#0001;  // new asynchronous result received
         #iprevMsgCounter := #IMsgCounter;  // store current value to detect the change
       END_REGION check for new result
     ELSE
       // on error replace values
       #XreMirrorbit := FALSE;
       #XreNewAsyncResult := FALSE;
     END_IF;  // on error replace values
   END_REGION read input data header of O3D3xx

   REGION set FB outputs
     IF #XErrorHW THEN  // invalid HW_ID
       #ErrorCodeFB := w#16#8100;  // error code for invalid HW_ID
     ELSE
       #ErrorCodeFB := w#16#0000;
     END_IF;
     #NewData := #XreMirrorbit OR #XreNewAsyncResult;  // new trigger response data
     IF #XreMirrorbit OR #XreNewAsyncResult THEN
       // transfer data into outputs
       #DIRdAddr := UDINT_TO_DINT(IN := #DIModuleInAddr + 12);  // set read address to first data Word
       #AllROIsGood := w#16#0001 = PEEK_WORD(area := 16#81, dbNumber := 0, byteOffset := #DIRdAddr);
       #DIRdAddr += 2;  // set read address to next Word
       IF #Tracking THEN
         // anchor tracking enabled
         #TrackingOK := w#16#0001 = PEEK_WORD(area := 16#81, dbNumber := 0, byteOffset := #DIRdAddr);
         #DIRdAddr += 2;  // set read address to next Word
       ELSE
         // anchor tracking disabled
         #TrackingOK := FALSE;
       END_IF;  // anchor tracking enabled

       FOR #IID := 0 TO 63 DO
         // initialize output values
         #ROI[#IID].Status := -1;
         #ROI[#IID].Value := -1;
       END_FOR;  // initialize output values

       #DILastRdAddr := UDINT_TO_DINT(IN := #DIModuleInAddr) + UINT_TO_DINT(#IModuleInLength - 6);  // calculate start address of last complete data set
       WHILE #DIRdAddr <= #DILastRdAddr DO
         // read ROI data
         #IID := WORD_TO_INT(PEEK_WORD(area := 16#81, dbNumber := 0, byteOffset := #DIRdAddr));  // read ROI ID
         IF #IID = 29556 THEN
           // value = "st" from end string "stop"
           EXIT;  // leave loop
         ELSE
           // end string not reached yet
           CASE #IID OF
             0..63:  // valid ID
               #ROI[#IID].Status := WORD_TO_INT(PEEK_WORD(area := 16#81, dbNumber := 0, byteOffset := #DIRdAddr + 2));  // copy statun into ROI
               #ROI[#IID].Value := WORD_TO_INT(PEEK_WORD(area := 16#81, dbNumber := 0, byteOffset := #DIRdAddr + 4));  // copy value into ROI
           END_CASE;
           #DIRdAddr += 6;  // set read address to next Word
         END_IF;  // end string not reached yet
       END_WHILE;  // read ROI data
     END_IF;  // transfer data into outputs
   END_REGION set FB outputs
END_FUNCTION_BLOCK

FUNCTION "ReadDataFn" : Void   // FC1, SCL
{ S7_Optimized_Access := 'TRUE' }
VERSION : 0.1
   VAR_INPUT
      TagPresent : Bool;
      Read : Bool;
   END_VAR
BEGIN
   IF #Read AND #TagPresent THEN
       "ReadData".RFIDValue :="TagValue";
       "ReadData".Object.Length :="O3D3xx_Dimensioning_DB".Length;
       "ReadData".Object.Width := "O3D3xx_Dimensioning_DB".Width ;
       "ReadData".Object.Height := "O3D3xx_Dimensioning_DB".Height ;
   END_IF;

   IF NOT #TagPresent THEN
       "ReadData".RFIDValue := 0;
       "ReadData".Object.Length := 0;
       "ReadData".Object.Width := 0;
       "ReadData".Object.Height := 0;
   END_IF;
END_FUNCTION

ORGANIZATION_BLOCK "Main"   // OB1, LAD, ProgramCycle
TITLE = "Main Program Sweep (Cycle)"
{ S7_Optimized_Access := 'TRUE' }
VERSION : 0.1
   VAR_INPUT
      Initial_Call : Bool;   // Initial call of this OB
      Remanence : Bool;   // =True, if remanent data are available
   END_VAR
   VAR_TEMP
      Scrap : UDInt;
      Trigger_Done : Bool;
   END_VAR
BEGIN

REGION Network 1: Trigger the O3D3xx sensor
   // Application 1 = my Dimensioning app
   // Application 2 = my Completeness app
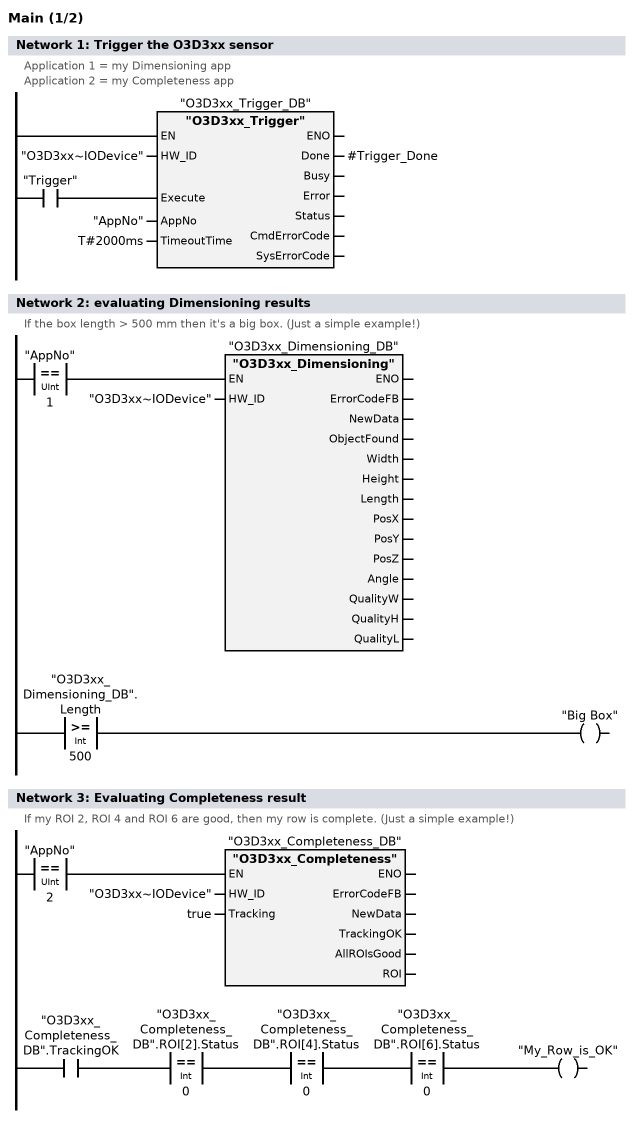
   RUNG wire#powerrail
      "O3D3xx_Trigger_DB"(Execute := wire#w1, HW_ID := "O3D3xx~IODevice", AppNo := "AppNo", TimeoutTime := T#2000ms, Done => #Trigger_Done, Busy =>, Error =>, Status =>, CmdErrorCode =>, SysErrorCode =>)
   END_RUNG
   RUNG wire#powerrail
      Contact( "Trigger" )
   END_RUNG wire#w1
   // the same network as SCL:
   "O3D3xx_Trigger_DB"(HW_ID := "O3D3xx~IODevice",   // "O3D3xx_Trigger"
                       Execute := "Trigger",
                       AppNo := "AppNo",
                       TimeoutTime := T#2000ms,
                       Done => #Trigger_Done);
END_REGION

REGION Network 2: evaluating Dimensioning results
   // If the box length > 500 mm then it's a big box. (Just a simple example!)
   RUNG wire#powerrail
      { S7_Templates := "SrcType := UInt" } EQ_Contact(in1 := "AppNo", in2 := 1)
      "O3D3xx_Dimensioning_DB"(HW_ID := "O3D3xx~IODevice", ErrorCodeFB =>, NewData =>, ObjectFound =>, Width =>, Height =>, Length =>, PosX =>, PosY =>, PosZ =>, Angle =>, QualityW =>, QualityH =>, QualityL =>)
   END_RUNG
   RUNG wire#powerrail
      { S7_Templates := "SrcType := Int" } GE_Contact(in1 := "O3D3xx_Dimensioning_DB".Length, in2 := 500)
      Coil( "Big Box" )
   END_RUNG
   // the same network as SCL:
   IF "AppNo" = 1 THEN
       "O3D3xx_Dimensioning_DB"(HW_ID := "O3D3xx~IODevice");   // "O3D3xx_Dimensioning"
   END_IF;
   "Big Box" := "O3D3xx_Dimensioning_DB".Length >= 500;
END_REGION

REGION Network 3: Evaluating Completeness result
   // If my ROI 2, ROI 4 and ROI 6 are good, then my row is complete. (Just a simple example!)
   RUNG wire#powerrail
      { S7_Templates := "SrcType := UInt" } EQ_Contact(in1 := "AppNo", in2 := 2)
      "O3D3xx_Completeness_DB"(HW_ID := "O3D3xx~IODevice", Tracking := true, ErrorCodeFB =>, NewData =>, TrackingOK =>, AllROIsGood =>, ROI =>)
   END_RUNG
   RUNG wire#powerrail
      Contact( "O3D3xx_Completeness_DB".TrackingOK )
      { S7_Templates := "SrcType := Int" } EQ_Contact(in1 := "O3D3xx_Completeness_DB".ROI[2].Status, in2 := 0)
      { S7_Templates := "SrcType := Int" } EQ_Contact(in1 := "O3D3xx_Completeness_DB".ROI[4].Status, in2 := 0)
      { S7_Templates := "SrcType := Int" } EQ_Contact(in1 := "O3D3xx_Completeness_DB".ROI[6].Status, in2 := 0)
      Coil( "My_Row_is_OK" )
   END_RUNG
   // the same network as SCL:
   IF "AppNo" = 2 THEN
       "O3D3xx_Completeness_DB"(HW_ID := "O3D3xx~IODevice", Tracking := true);   // "O3D3xx_Completeness"
   END_IF;
   "My_Row_is_OK" := "O3D3xx_Completeness_DB".TrackingOK AND ("O3D3xx_Completeness_DB".ROI[2].Status = 0) AND ("O3D3xx_Completeness_DB".ROI[4].Status = 0) AND ("O3D3xx_Completeness_DB".ROI[6].Status = 0);
END_REGION

REGION Network 4: Get scrap rate
   // Just a simple example!
   // After each trigger it reads the statistics. If the FAIL rate is more than 3% it triggers an alarm.
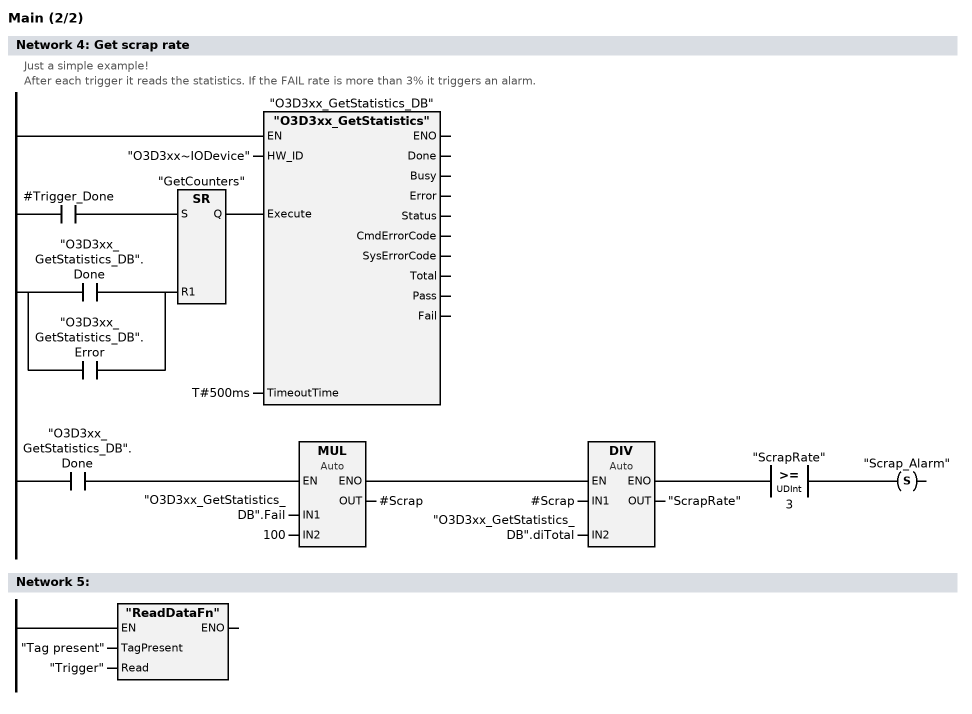
   RUNG wire#powerrail
      "O3D3xx_GetStatistics_DB"(Execute := wire#w2, HW_ID := "O3D3xx~IODevice", TimeoutTime := T#500ms, Done =>, Busy =>, Error =>, Status =>, CmdErrorCode =>, SysErrorCode =>, Total =>, Pass =>, Fail =>)
   END_RUNG
   RUNG wire#powerrail
      Contact( #Trigger_Done )
      S_SR(operand := "GetCounters", r1 := wire#w1)
   END_RUNG wire#w2
   RUNG wire#powerrail
      Contact( "O3D3xx_GetStatistics_DB".Done )
   END_RUNG wire#w1
   RUNG wire#powerrail
      Contact( "O3D3xx_GetStatistics_DB".Error )
   END_RUNG wire#w1
   RUNG wire#powerrail
      Contact( "O3D3xx_GetStatistics_DB".Done )
      Mul(in1 := "O3D3xx_GetStatistics_DB".Fail, in2 := 100, out => #Scrap)
      Div(in1 := #Scrap, in2 := "O3D3xx_GetStatistics_DB".diTotal, out => "ScrapRate")
      { S7_Templates := "SrcType := UDInt" } GE_Contact(in1 := "ScrapRate", in2 := 3)
      S_Coil( "Scrap_Alarm" )
   END_RUNG
   // the same network as SCL:
   IF #Trigger_Done THEN
       "GetCounters" := TRUE;   // SR flip-flop
   END_IF;
   IF "O3D3xx_GetStatistics_DB".Done OR "O3D3xx_GetStatistics_DB".Error THEN "GetCounters" := FALSE; END_IF;
   "O3D3xx_GetStatistics_DB"(HW_ID := "O3D3xx~IODevice", Execute := "GetCounters", TimeoutTime := T#500ms);   // "O3D3xx_GetStatistics"
   IF "O3D3xx_GetStatistics_DB".Done THEN
       #Scrap := "O3D3xx_GetStatistics_DB".Fail * 100;
       "ScrapRate" := #Scrap / "O3D3xx_GetStatistics_DB".diTotal;
   END_IF;
   IF "O3D3xx_GetStatistics_DB".Done AND ("ScrapRate" >= 3) THEN "Scrap_Alarm" := TRUE; END_IF;
END_REGION

REGION Network 5
   RUNG wire#powerrail
      "ReadDataFn"(TagPresent := "Tag present", Read := "Trigger")
   END_RUNG
   // the same network as SCL:
   "ReadDataFn"(TagPresent := "Tag present", Read := "Trigger");
END_REGION
END_ORGANIZATION_BLOCK

(* ===== HMI "HMI_RT_1" =====
system functions are stored by id; their names below are inferred from use
connection "HMI_Connection_1": ETHERNET, S7_1200_OMS

HMI tags "Default tag table"
   "Tag_ScreenNumber" : UInt, internal
   "Trigger" : Bool = PLC Trigger AT %M0.0, 1 s
   "O3D3xx_Dimensioning_DB_Length" : Int = PLC O3D3xx_Dimensioning_DB.Length, 1 s
   "O3D3xx_Dimensioning_DB_Width" : Int = PLC O3D3xx_Dimensioning_DB.Width, 1 s
   "O3D3xx_Dimensioning_DB_Height" : Int = PLC O3D3xx_Dimensioning_DB.Height, 1 s
   "Tag present" : Bool = PLC "Tag present" AT %I519.2, 1 s
   "TagValue" : Byte = PLC TagValue AT %IB520, 1 s
   "ReadData_RFIDValue" : Byte = PLC ReadData.RFIDValue, 1 s
   "ReadData_Object_Length" : Int = PLC ReadData.Object.Length, 1 s
   "ReadData_Object_Width" : Int = PLC ReadData.Object.Width, 1 s
   "ReadData_Object_Height" : Int = PLC ReadData.Object.Height, 1 s

screen "Root screen" 800x420, template "Template_1"
   on GenerateScreen: SetTag("Tag_ScreenNumber", 1)
   Button "Button_1" at 111,189 size 211x53; TextOff 'READ VALUE'
      on Press: function_b14e0dd5("Trigger", 0)
      Appearance <- "Trigger"
   IOField "I/O field_1" at 651,135 size 56x45; FormatPattern 999
      ProcessValue <- "ReadData_RFIDValue"
   IOField "I/O field_2" at 651,193 size 57x45; FormatPattern 999
      ProcessValue <- "ReadData_Object_Length"
   IOField "I/O field_3" at 651,255 size 57x45; FormatPattern 999
      ProcessValue <- "ReadData_Object_Width"
   IOField "I/O field_4" at 651,317 size 57x45; FormatPattern 999
      ProcessValue <- "ReadData_Object_Height"
   TextField "Text field_1" at 492,137 size 137x37; Text 'RFID Value'
   TextField "Text field_2" at 545,199 size 86x37; Text 'Length'
   TextField "Text field_3" at 558,260 size 74x37; Text 'Width'
   TextField "Text field_4" at 548,320 size 82x37; Text 'Height'
   TextField "Text field_5" at 8,13 size 782x33; Text 'IFM RFID and 3D Camera Integration with Siemens S7-1200'
   Rectangle "Rectangle_2" at 113,145 size 25x21
      Appearance <- "Tag present"
   TextField "Text field_6" at 147,136 size 160x37; Text 'Tag detected'
   TextField "Text field_7" at 421,85 size 342x37; Text 'OBJECT INFORMATION'
   TextField "Text field_8" at 50,86 size 288x37; Text 'TRIGGER CONTROL'

Template "Template_1" 800x420
   Button "Exit" at 720,360 size 78x58; TextOff 'Exit'; PictureOff "ExitRuntime_TP700_Comfort_TR"; PictureOn "ExitRuntime_TP700_Comfort_TR"
      on Release: StopRuntime(0)
*)